FUNCTION_BLOCK DLG_MessageBox (* VT-Dialog wie Windows-MessageBox (eine Instanz je Anwendung) *)
  (* Standard: 61499-2; Description: Copyright (c) 2026 Meisterschulen am Ostbahnhof This program and the accompanying materials are made available under the terms of the Eclipse Public License 2.0 which is available at https://www.eclipse.org/legal/epl-2.0/ SPDX-License-Identifier: EPL-2.0 *)
  (* Version 1.1, 2026-11-25, Franz Höpfinger, Meisterschulen am Ostbahnhof, SubApp -> Composite FB (Lib wird wegen DLG_CTRL ohnehin gebaut, im fboot nur eine Instanz). *)
  (* Version 1.0, 2026-11-17, Franz Höpfinger, Meisterschulen am Ostbahnhof, initial API and implementation and/or initial documentation *)
  PACKAGE isobus::UT::dialog;
  IMPORT isobus::UT::Q::const::IDs::ID_NULL;
  IMPORT isobus::UT::dialog::DialogIDs::Button_Dlg_Abort;
  IMPORT isobus::UT::dialog::DialogIDs::Button_Dlg_Cancel;
  IMPORT isobus::UT::dialog::DialogIDs::Button_Dlg_Ignore;
  IMPORT isobus::UT::dialog::DialogIDs::Button_Dlg_No;
  IMPORT isobus::UT::dialog::DialogIDs::Button_Dlg_OK;
  IMPORT isobus::UT::dialog::DialogIDs::Button_Dlg_Retry;
  IMPORT isobus::UT::dialog::DialogIDs::Button_Dlg_Yes;
  IMPORT isobus::UT::dialog::DialogIDs::Container_Dialog;
  IMPORT isobus::UT::dialog::DialogIDs::FillAttributes_Dlg_Title;
  IMPORT isobus::UT::dialog::DialogIDs::ObjectPointer_Dlg_Buttons;
  IMPORT isobus::UT::dialog::DialogIDs::ObjectPointer_Dlg_Cover;
  IMPORT isobus::UT::dialog::DialogIDs::ObjectPointer_Dlg_Icon;
  IMPORT isobus::UT::dialog::DialogIDs::ObjectPointer_Dlg_Text;
  IMPORT isobus::UT::dialog::DialogIDs::ObjectPointer_Dlg_Title;
  IMPORT isobus::UT::io::Button::ButtonActivationCode::BT_RELEASED_UNLATCHED;
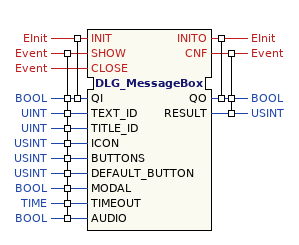
  EVENT_INPUT
    INIT : EInit WITH QI; (* Initialisierung *)
    SHOW WITH QI, TEXT_ID, TITLE_ID, ICON, BUTTONS, DEFAULT_BUTTON, MODAL, TIMEOUT, AUDIO; (* Dialog zeigen *)
    CLOSE; (* Dialog schliessen *)
  END_EVENT
  EVENT_OUTPUT
    INITO : EInit WITH QO; (* Initialisierung fertig *)
    CNF WITH QO, RESULT; (* Dialog beendet, RESULT gueltig *)
  END_EVENT
  VAR_INPUT
    QI : BOOL := TRUE; (* Freigabe *)
    TEXT_ID : UINT := ID_NULL; (* OutputString Meldungstext *)
    TITLE_ID : UINT := ID_NULL; (* OutputString Titel, NULL = Standard je Icon *)
    ICON : USINT := USINT#1; (* DLG_ICON_* *)
    BUTTONS : USINT := USINT#1; (* DLG_BTN_* *)
    DEFAULT_BUTTON : USINT := USINT#1; (* Fokus auf Taste 1..3 *)
    MODAL : BOOL := FALSE; (* Maske abdecken *)
    TIMEOUT : TIME := T#0s; (* T#0s = kein Timeout *)
    AUDIO : BOOL := FALSE; (* Ton beim Oeffnen *)
  END_VAR
  VAR_OUTPUT
    QO : BOOL; (* Qualitaet *)
    RESULT : USINT; (* DLG_RES_* *)
  END_VAR
  FBS
    CTRL : isobus::UT::dialog::DLG_CTRL;
    QN_COVER : isobus::UT::Q::Q_NumericValue(QI := TRUE, u16ObjId := ObjectPointer_Dlg_Cover);
    QN_ICON : isobus::UT::Q::Q_NumericValue(QI := TRUE, u16ObjId := ObjectPointer_Dlg_Icon);
    QN_TITLE : isobus::UT::Q::Q_NumericValue(QI := TRUE, u16ObjId := ObjectPointer_Dlg_Title);
    QN_TEXT : isobus::UT::Q::Q_NumericValue(QI := TRUE, u16ObjId := ObjectPointer_Dlg_Text);
    QN_BUTTONS : isobus::UT::Q::Q_NumericValue(QI := TRUE, u16ObjId := ObjectPointer_Dlg_Buttons);
    QF_TITLE : isobus::UT::Q::Q_FillAttributes(QI := TRUE, u16ObjId := FillAttributes_Dlg_Title, u8FillType := USINT#2, u16FillPatternId := ID_NULL);
    QH_SHOW : isobus::UT::Q::Q_ObjHideShow(QI := TRUE, u16ObjId := Container_Dialog, qVisible := BYTE#1);
    QH_HIDE : isobus::UT::Q::Q_ObjHideShow(QI := TRUE, u16ObjId := Container_Dialog, qVisible := BYTE#0);
    FOCUS : iec61499::events::E_DEMUX_8;
    QS_OK : isobus::UT::Q::Q_ObjSelectInput(QI := TRUE, u16ObjId := Button_Dlg_OK, u8Option := USINT#255);
    QS_CANCEL : isobus::UT::Q::Q_ObjSelectInput(QI := TRUE, u16ObjId := Button_Dlg_Cancel, u8Option := USINT#255);
    QS_ABORT : isobus::UT::Q::Q_ObjSelectInput(QI := TRUE, u16ObjId := Button_Dlg_Abort, u8Option := USINT#255);
    QS_RETRY : isobus::UT::Q::Q_ObjSelectInput(QI := TRUE, u16ObjId := Button_Dlg_Retry, u8Option := USINT#255);
    QS_IGNORE : isobus::UT::Q::Q_ObjSelectInput(QI := TRUE, u16ObjId := Button_Dlg_Ignore, u8Option := USINT#255);
    QS_YES : isobus::UT::Q::Q_ObjSelectInput(QI := TRUE, u16ObjId := Button_Dlg_Yes, u8Option := USINT#255);
    QS_NO : isobus::UT::Q::Q_ObjSelectInput(QI := TRUE, u16ObjId := Button_Dlg_No, u8Option := USINT#255);
    FOCUS_DONE : iec61499::events::E_MUX_8;
    AUDIO_SW : iec61499::events::E_SWITCH;
    Q_AUDIO : isobus::UT::Q::Q_CtrlAudioSignal(QI := TRUE, u8NumOfRepit := USINT#1, u16Frequency := UINT#2000, u16OnTimeMs := UINT#100, u16OffTimeMs := UINT#0);
    AUDIO_DONE : iec61499::events::E_MERGE;
    TIMER : iec61499::events::E_DELAY;
    BTN_OK : isobus::UT::io::Button::Button_IE(QI := TRUE, u16ObjId := Button_Dlg_OK, InputEvent := BT_RELEASED_UNLATCHED);
    BTN_CANCEL : isobus::UT::io::Button::Button_IE(QI := TRUE, u16ObjId := Button_Dlg_Cancel, InputEvent := BT_RELEASED_UNLATCHED);
    BTN_ABORT : isobus::UT::io::Button::Button_IE(QI := TRUE, u16ObjId := Button_Dlg_Abort, InputEvent := BT_RELEASED_UNLATCHED);
    BTN_RETRY : isobus::UT::io::Button::Button_IE(QI := TRUE, u16ObjId := Button_Dlg_Retry, InputEvent := BT_RELEASED_UNLATCHED);
    BTN_IGNORE : isobus::UT::io::Button::Button_IE(QI := TRUE, u16ObjId := Button_Dlg_Ignore, InputEvent := BT_RELEASED_UNLATCHED);
    BTN_YES : isobus::UT::io::Button::Button_IE(QI := TRUE, u16ObjId := Button_Dlg_Yes, InputEvent := BT_RELEASED_UNLATCHED);
    BTN_NO : isobus::UT::io::Button::Button_IE(QI := TRUE, u16ObjId := Button_Dlg_No, InputEvent := BT_RELEASED_UNLATCHED);
  END_FBS
  EVENT_CONNECTIONS
    BTN_OK.IND TO CTRL.B_OK;
    BTN_CANCEL.IND TO CTRL.B_CANCEL;
    BTN_ABORT.IND TO CTRL.B_ABORT;
    BTN_RETRY.IND TO CTRL.B_RETRY;
    BTN_IGNORE.IND TO CTRL.B_IGNORE;
    BTN_YES.IND TO CTRL.B_YES;
    BTN_NO.IND TO CTRL.B_NO;
    CTRL.SHOWO TO QN_COVER.REQ;
    QN_COVER.CNF TO QN_ICON.REQ;
    QN_ICON.CNF TO QN_TITLE.REQ;
    QN_TITLE.CNF TO QN_TEXT.REQ;
    QN_TEXT.CNF TO QN_BUTTONS.REQ;
    QN_BUTTONS.CNF TO QF_TITLE.REQ;
    QF_TITLE.CNF TO QH_SHOW.REQ;
    QH_SHOW.CNF TO FOCUS.EI;
    FOCUS.EO1 TO QS_OK.REQ;
    QS_OK.CNF TO FOCUS_DONE.EI1;
    FOCUS.EO2 TO QS_CANCEL.REQ;
    QS_CANCEL.CNF TO FOCUS_DONE.EI2;
    FOCUS.EO3 TO QS_ABORT.REQ;
    QS_ABORT.CNF TO FOCUS_DONE.EI3;
    FOCUS.EO4 TO QS_RETRY.REQ;
    QS_RETRY.CNF TO FOCUS_DONE.EI4;
    FOCUS.EO5 TO QS_IGNORE.REQ;
    QS_IGNORE.CNF TO FOCUS_DONE.EI5;
    FOCUS.EO6 TO QS_YES.REQ;
    QS_YES.CNF TO FOCUS_DONE.EI6;
    FOCUS.EO7 TO QS_NO.REQ;
    QS_NO.CNF TO FOCUS_DONE.EI7;
    FOCUS.EO8 TO FOCUS_DONE.EI8;
    FOCUS_DONE.EO TO AUDIO_SW.EI;
    AUDIO_SW.EO0 TO AUDIO_DONE.EI1;
    AUDIO_SW.EO1 TO Q_AUDIO.REQ;
    Q_AUDIO.CNF TO AUDIO_DONE.EI2;
    AUDIO_DONE.EO TO CTRL.SHOWN;
    CTRL.HIDEO TO QH_HIDE.REQ;
    QH_HIDE.CNF TO CTRL.HIDDEN;
    CTRL.START_T TO TIMER.START;
    CTRL.STOP_T TO TIMER.STOP;
    TIMER.EO TO CTRL.TMO;
    INIT TO BTN_OK.INIT;
    CTRL.INITO TO QN_COVER.INIT;
    QN_COVER.INITO TO QN_ICON.INIT;
    QN_ICON.INITO TO QN_TITLE.INIT;
    QN_TITLE.INITO TO QN_TEXT.INIT;
    QN_TEXT.INITO TO QN_BUTTONS.INIT;
    QN_BUTTONS.INITO TO QF_TITLE.INIT;
    QF_TITLE.INITO TO QH_SHOW.INIT;
    QH_SHOW.INITO TO QH_HIDE.INIT;
    QH_HIDE.INITO TO QS_OK.INIT;
    QS_OK.INITO TO QS_CANCEL.INIT;
    QS_CANCEL.INITO TO QS_ABORT.INIT;
    QS_ABORT.INITO TO QS_RETRY.INIT;
    QS_RETRY.INITO TO QS_IGNORE.INIT;
    QS_IGNORE.INITO TO QS_YES.INIT;
    QS_YES.INITO TO QS_NO.INIT;
    QS_NO.INITO TO Q_AUDIO.INIT;
    BTN_OK.INITO TO BTN_CANCEL.INIT;
    BTN_CANCEL.INITO TO BTN_ABORT.INIT;
    BTN_ABORT.INITO TO BTN_RETRY.INIT;
    BTN_RETRY.INITO TO BTN_IGNORE.INIT;
    BTN_IGNORE.INITO TO BTN_YES.INIT;
    BTN_YES.INITO TO BTN_NO.INIT;
    SHOW TO CTRL.SHOW;
    CLOSE TO CTRL.CLOSE;
    CTRL.CNF TO CNF;
    BTN_NO.INITO TO CTRL.INIT;
    Q_AUDIO.INITO TO INITO;
  END_CONNECTIONS
  DATA_CONNECTIONS
    CTRL.COVER_ID TO QN_COVER.u32NewValue;
    CTRL.ICON_ID TO QN_ICON.u32NewValue;
    CTRL.TITLE_ID_O TO QN_TITLE.u32NewValue;
    CTRL.TEXT_ID_O TO QN_TEXT.u32NewValue;
    CTRL.BUTTONS_ID TO QN_BUTTONS.u32NewValue;
    CTRL.TITLE_COLOUR TO QF_TITLE.u8FillColour;
    CTRL.FOCUS_K TO FOCUS.K;
    CTRL.AUDIO_O TO AUDIO_SW.G;
    CTRL.TIMEOUT_O TO TIMER.DT;
    QI TO CTRL.QI;
    TEXT_ID TO CTRL.TEXT_ID;
    TITLE_ID TO CTRL.TITLE_ID;
    ICON TO CTRL.ICON;
    BUTTONS TO CTRL.BUTTONS;
    DEFAULT_BUTTON TO CTRL.DEFAULT_BUTTON;
    MODAL TO CTRL.MODAL;
    TIMEOUT TO CTRL.TIMEOUT;
    AUDIO TO CTRL.AUDIO;
    CTRL.QO TO QO;
    CTRL.RESULT TO RESULT;
  END_CONNECTIONS
END_FUNCTION_BLOCK
